// TIA Portal V20 export
FUNCTION_BLOCK "Main_Safety_RTG1"   // FB3, F_LAD
{ S7_Optimized_Access := 'TRUE' }
// stored: AutoNumber false
   VAR
      "ESTOP1_NOT-HALT Taster1" : ESTOP1;
      "stat_Q_NOT-HALT Taster1" : Bool;
      "stat_AckReq_NOT-HALT Taster1" : Bool;
      "ESTOP1_NOT-HALT Extern 1" : ESTOP1;
      "stat_Q_NOT-HALT Extern 1" : Bool;
      "stat_AckReq_NOT-HALT Extern1" : Bool;
      "ESTOP1_NOT-HALT Extern 2" : ESTOP1;
      "stat_Q_NOT-HALT Extern 2" : Bool;
      "stat_AckReq_NOT-HALT Extern 2" : Bool;
      "ESTOP1_Tür 1" : ESTOP1;
      "stat_Q_Tür 1" : Bool;
      "stat_AckReq_Tür 1" : Bool;
      "ESTOP1_Tür 2" : ESTOP1;
      "stat_Q_Tür 2" : Bool;
      "stat_AckReq_Tür 2" : Bool;
      ESTOP1_Systemdruck : ESTOP1;
      stat_AckReq_Systemdruck : Bool;
      "FDBACK_1_NOT-HALT Schütz mit DE_NOT-HALT_Schuetz_Rueckf" : FDBACK;
      "stat_Q_FDBK_1_NOT-HALT Schütz mit DE_NOT-HALT_Schuetz_Rueckf" : Bool;
      "stat_ERROR_FDBK_1_NOT-HALT Schütz mit DE_NOT-HALT_Schuetz_Rueckf" : Bool;
      "FDBACK_2_NOT-HALT Schütz mit IS_Rueck_Entlueftung" : FDBACK;
      "stat_Q_FDBK_2_NOT-HALT Schütz mit IS_Rueck_Entlueftung" : Bool;
      "stat_ERROR_FDBK_2_NOT-HALT Schütz mit IS_Rueck_Entlueftung" : Bool;
      "FDBACK_3_NOT-HALT Schütz mit IS_Druckbereich_entlueftet" : FDBACK;
      "stat_Q_FDBK_3_NOT-HALT Schütz mit IS_Druckbereich_entlueftet" : Bool;
      "stat_ERROR_FDBK_3_NOT-HALT Schütz mit IS_Druckbereich_entlueftet" : Bool;
      "FDBACK_4_NOT-HALT Türe 1 RST mit DE_NOT-HALT_Tuere_1_Rueck_RST" : FDBACK;
      "stat_Q_FDBK_4_NOT-HALT Türe 1 RST mit DE_NOT-HALT_Tuere_1_Rueck_RST" : Bool;
      "stat_ERROR_FDBK_4_NOT-HALT Türe 1 RST mit DE_NOT-HALT_Tuere_1_Rueck_RST" : Bool;
      "FDBACK_5_NOT-HALT Türe 1 mit DE_NOT-HALT_Tuere_1_Rueckf" : FDBACK;
      "stat_Q_FDBK_5_NOT-HALT Türe 1 mit DE_NOT-HALT_Tuere_1_Rueckf" : Bool;
      "stat_ERROR_FDBK_5_NOT-HALT Türe 1 mit DE_NOT-HALT_Tuere_1_Rueckf" : Bool;
      "FDBACK_6_NOT-HALT Türe 1 mit DE_Antriebe_Rueckf" : FDBACK;
      "stat_Q_FDBK_6_NOT-HALT Türe 1 mit DE_Antriebe_Rueckf" : Bool;
      "stat_ERROR_FDBK_6_NOT-HALT Türe 1 mit DE_Antriebe_Rueckf" : Bool;
      "FDBACK_7_NOT-HALT Türe 2 RST mit DE_NOT-HALT_Tuere_2_Rueck_RST" : FDBACK;
      "stat_Q_FDBK_7_NOT-HALT Türe 2 RST mit DE_NOT-HALT_Tuere_2_Rueck_RST" : Bool;
      "stat_ERROR_FDBK_7_NOT-HALT Türe 2 RST mit DE_NOT-HALT_Tuere_2_Rueck_RST" : Bool;
      "FDBACK_8_NOT-HALT Türe 2 mit DE_NOT-HALT_Tuere_2_Rueckf" : FDBACK;
      "stat_Q_FDBK_8_NOT-HALT Türe 2 mit DE_NOT-HALT_Tuere_2_Rueckf" : Bool;
      "stat_ERROR_FDBK_8_NOT-HALT Türe 2 mit DE_NOT-HALT_Tuere_2_Rueckf" : Bool;
      "FDBACK_10_Sicherere Bewegung" : FDBACK;
      "stat_AckReq_10_Sicherere Bewegung" : Bool;
      ACK_GL_Instance : ACK_GL;
      Systemdruck_OK : Bool;
      Antriebe_sicher : Bool;
      "TON_Zuhaltung_Freigben_mit_NOT-HALT" : TON;
      BA_0_groesser_1_5 : Bool;
      TON_BA_0_groesser_1_5 : TON;
      TON_Türen_setzen_zum_öffnen : TON;
      BA_0 : Bool;
      Zuhaltung_freigegeben : Bool;
   END_VAR
BEGIN

REGION Network 1: IS100_0/IS101_0 (2v2) NOT-HALT Taster 1
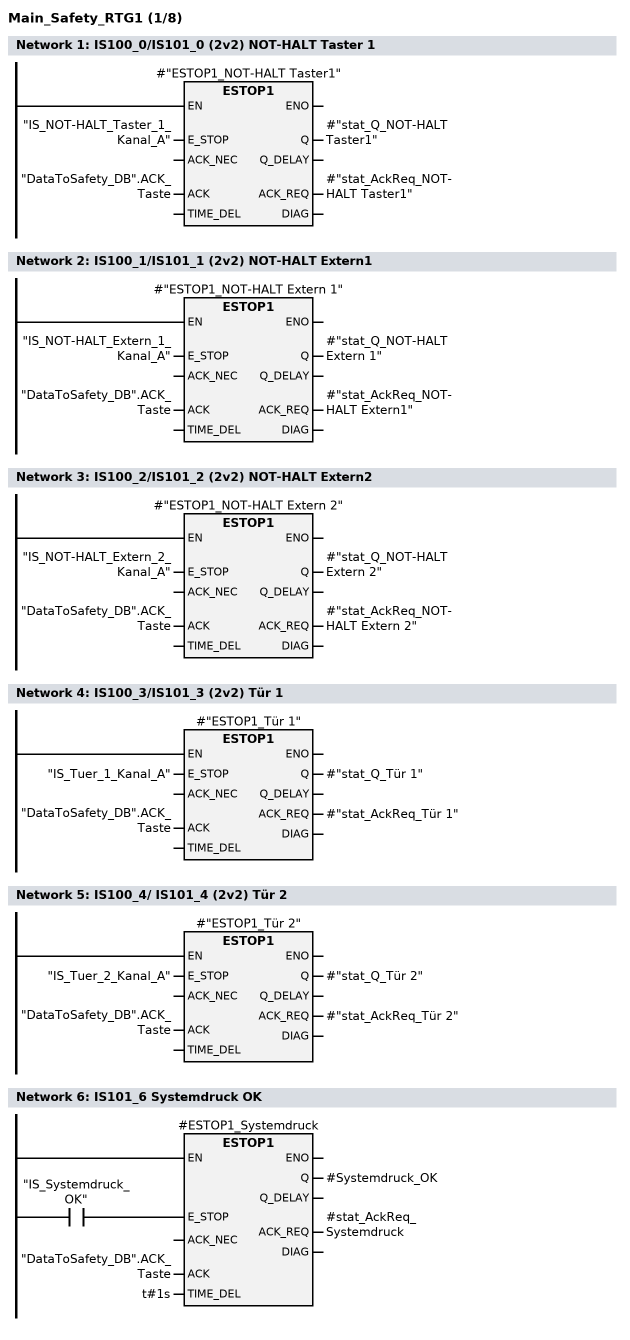
   RUNG wire#powerrail
      #"ESTOP1_NOT-HALT Taster1".ESTOP1(E_STOP := "IS_NOT-HALT_Taster_1_Kanal_A", ACK_NEC :=, ACK := "DataToSafety_DB".ACK_Taste, TIME_DEL :=, Q => #"stat_Q_NOT-HALT Taster1", Q_DELAY =>, ACK_REQ => #"stat_AckReq_NOT-HALT Taster1", DIAG =>)
   END_RUNG
   // the same network as SCL:
   #"ESTOP1_NOT-HALT Taster1"(E_STOP := "IS_NOT-HALT_Taster_1_Kanal_A",   // ESTOP1
                           ACK := "DataToSafety_DB".ACK_Taste,
                           Q => #"stat_Q_NOT-HALT Taster1",
                           ACK_REQ => #"stat_AckReq_NOT-HALT Taster1");
END_REGION

REGION Network 2: IS100_1/IS101_1 (2v2) NOT-HALT Extern1
   RUNG wire#powerrail
      #"ESTOP1_NOT-HALT Extern 1".ESTOP1(E_STOP := "IS_NOT-HALT_Extern_1_Kanal_A", ACK_NEC :=, ACK := "DataToSafety_DB".ACK_Taste, TIME_DEL :=, Q => #"stat_Q_NOT-HALT Extern 1", Q_DELAY =>, ACK_REQ => #"stat_AckReq_NOT-HALT Extern1", DIAG =>)
   END_RUNG
   // the same network as SCL:
   #"ESTOP1_NOT-HALT Extern 1"(E_STOP := "IS_NOT-HALT_Extern_1_Kanal_A",   // ESTOP1
                           ACK := "DataToSafety_DB".ACK_Taste,
                           Q => #"stat_Q_NOT-HALT Extern 1",
                           ACK_REQ => #"stat_AckReq_NOT-HALT Extern1");
END_REGION

REGION Network 3: IS100_2/IS101_2 (2v2) NOT-HALT Extern2
   RUNG wire#powerrail
      #"ESTOP1_NOT-HALT Extern 2".ESTOP1(E_STOP := "IS_NOT-HALT_Extern_2_Kanal_A", ACK_NEC :=, ACK := "DataToSafety_DB".ACK_Taste, TIME_DEL :=, Q => #"stat_Q_NOT-HALT Extern 2", Q_DELAY =>, ACK_REQ => #"stat_AckReq_NOT-HALT Extern 2", DIAG =>)
   END_RUNG
   // the same network as SCL:
   #"ESTOP1_NOT-HALT Extern 2"(E_STOP := "IS_NOT-HALT_Extern_2_Kanal_A",   // ESTOP1
                           ACK := "DataToSafety_DB".ACK_Taste,
                           Q => #"stat_Q_NOT-HALT Extern 2",
                           ACK_REQ => #"stat_AckReq_NOT-HALT Extern 2");
END_REGION

REGION Network 4: IS100_3/IS101_3 (2v2) Tür 1
   RUNG wire#powerrail
      #"ESTOP1_Tür 1".ESTOP1(E_STOP := "IS_Tuer_1_Kanal_A", ACK_NEC :=, ACK := "DataToSafety_DB".ACK_Taste, TIME_DEL :=, Q => #"stat_Q_Tür 1", Q_DELAY =>, ACK_REQ => #"stat_AckReq_Tür 1", DIAG =>)
   END_RUNG
   // the same network as SCL:
   #"ESTOP1_Tür 1"(E_STOP := "IS_Tuer_1_Kanal_A",   // ESTOP1
                   ACK := "DataToSafety_DB".ACK_Taste,
                   Q => #"stat_Q_Tür 1",
                   ACK_REQ => #"stat_AckReq_Tür 1");
END_REGION

REGION Network 5: IS100_4/ IS101_4 (2v2) Tür 2
   RUNG wire#powerrail
      #"ESTOP1_Tür 2".ESTOP1(E_STOP := "IS_Tuer_2_Kanal_A", ACK_NEC :=, ACK := "DataToSafety_DB".ACK_Taste, TIME_DEL :=, Q => #"stat_Q_Tür 2", Q_DELAY =>, ACK_REQ => #"stat_AckReq_Tür 2", DIAG =>)
   END_RUNG
   // the same network as SCL:
   #"ESTOP1_Tür 2"(E_STOP := "IS_Tuer_2_Kanal_A",   // ESTOP1
                   ACK := "DataToSafety_DB".ACK_Taste,
                   Q => #"stat_Q_Tür 2",
                   ACK_REQ => #"stat_AckReq_Tür 2");
END_REGION

REGION Network 6: IS101_6 Systemdruck OK
   RUNG wire#powerrail
      #ESTOP1_Systemdruck.ESTOP1(E_STOP := wire#w1, ACK_NEC :=, ACK := "DataToSafety_DB".ACK_Taste, TIME_DEL := t#1s, Q => #Systemdruck_OK, Q_DELAY =>, ACK_REQ => #stat_AckReq_Systemdruck, DIAG =>)
   END_RUNG
   RUNG wire#powerrail
      Contact( "IS_Systemdruck_OK" )
   END_RUNG wire#w1
   // the same network as SCL:
   #ESTOP1_Systemdruck(E_STOP := "IS_Systemdruck_OK",   // ESTOP1
                       ACK := "DataToSafety_DB".ACK_Taste,
                       TIME_DEL := t#1s,
                       Q => #Systemdruck_OK,
                       ACK_REQ => #stat_AckReq_Systemdruck);
END_REGION

REGION Network 7: Antriebe sicher
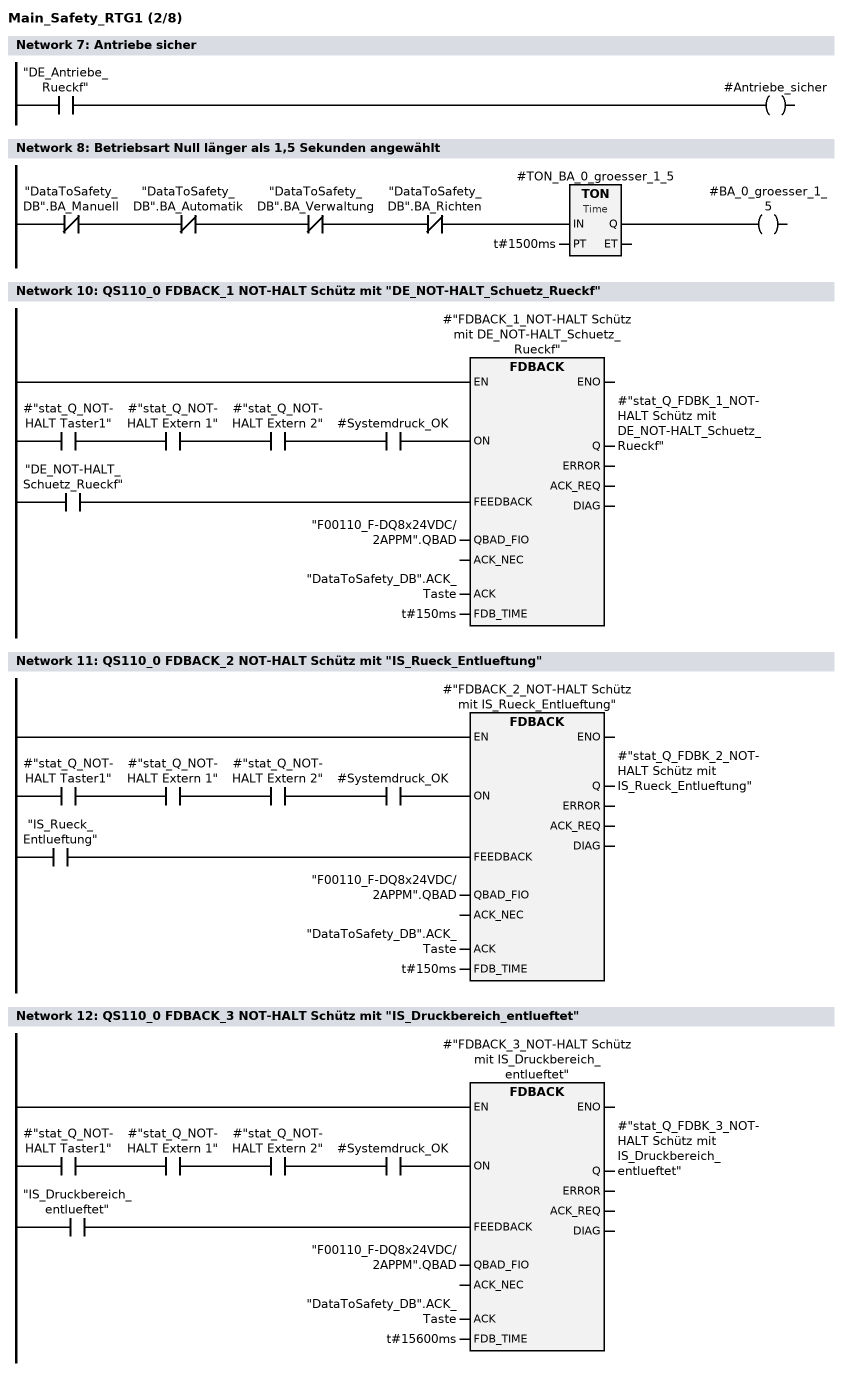
   RUNG wire#powerrail
      Contact( "DE_Antriebe_Rueckf" )
      Coil( #Antriebe_sicher )
   END_RUNG
   // the same network as SCL:
   #Antriebe_sicher := "DE_Antriebe_Rueckf";
END_REGION

REGION Network 8: Betriebsart Null länger als 1,5 Sekunden angewählt
   RUNG wire#powerrail
      I_Contact( "DataToSafety_DB".BA_Manuell )
      I_Contact( "DataToSafety_DB".BA_Automatik )
      I_Contact( "DataToSafety_DB".BA_Verwaltung )
      I_Contact( "DataToSafety_DB".BA_Richten )
      { S7_Templates := "[time_type := Time, codedbool_type := DInt]" } #TON_BA_0_groesser_1_5.TON(pt := t#1500ms, et =>)
      Coil( #BA_0_groesser_1_5 )
   END_RUNG
   // the same network as SCL:
   #TON_BA_0_groesser_1_5.TON(IN := NOT "DataToSafety_DB".BA_Manuell AND NOT "DataToSafety_DB".BA_Automatik AND NOT "DataToSafety_DB".BA_Verwaltung AND NOT "DataToSafety_DB".BA_Richten,
                           PT := t#1500ms);
   #BA_0_groesser_1_5 := #TON_BA_0_groesser_1_5.Q;
END_REGION

REGION Network 9: *********************************************************************************************
END_REGION

REGION Network 10: QS110_0 FDBACK_1 NOT-HALT Schütz mit "DE_NOT-HALT_Schuetz_Rueckf"
   RUNG wire#powerrail
      #"FDBACK_1_NOT-HALT Schütz mit DE_NOT-HALT_Schuetz_Rueckf".FDBACK(ON := wire#w1, FEEDBACK := wire#w2, QBAD_FIO := "F00110_F-DQ8x24VDC/2APPM".QBAD, ACK_NEC :=, ACK := "DataToSafety_DB".ACK_Taste, FDB_TIME := t#150ms, Q => #"stat_Q_FDBK_1_NOT-HALT Schütz mit DE_NOT-HALT_Schuetz_Rueckf", ERROR =>, ACK_REQ =>, DIAG =>)
   END_RUNG
   RUNG wire#powerrail
      Contact( #"stat_Q_NOT-HALT Taster1" )
      Contact( #"stat_Q_NOT-HALT Extern 1" )
      Contact( #"stat_Q_NOT-HALT Extern 2" )
      Contact( #Systemdruck_OK )
   END_RUNG wire#w1
   RUNG wire#powerrail
      Contact( "DE_NOT-HALT_Schuetz_Rueckf" )
   END_RUNG wire#w2
   // the same network as SCL:
   #"FDBACK_1_NOT-HALT Schütz mit DE_NOT-HALT_Schuetz_Rueckf"(ON := #"stat_Q_NOT-HALT Taster1" AND #"stat_Q_NOT-HALT Extern 1" AND #"stat_Q_NOT-HALT Extern 2" AND #Systemdruck_OK,   // FDBACK
                           FEEDBACK := "DE_NOT-HALT_Schuetz_Rueckf",
                           QBAD_FIO := "F00110_F-DQ8x24VDC/2APPM".QBAD,
                           ACK := "DataToSafety_DB".ACK_Taste,
                           FDB_TIME := t#150ms,
                           Q => #"stat_Q_FDBK_1_NOT-HALT Schütz mit DE_NOT-HALT_Schuetz_Rueckf");
END_REGION

REGION Network 11: QS110_0 FDBACK_2 NOT-HALT Schütz mit "IS_Rueck_Entlueftung"
   RUNG wire#powerrail
      #"FDBACK_2_NOT-HALT Schütz mit IS_Rueck_Entlueftung".FDBACK(ON := wire#w1, FEEDBACK := wire#w2, QBAD_FIO := "F00110_F-DQ8x24VDC/2APPM".QBAD, ACK_NEC :=, ACK := "DataToSafety_DB".ACK_Taste, FDB_TIME := t#150ms, Q => #"stat_Q_FDBK_2_NOT-HALT Schütz mit IS_Rueck_Entlueftung", ERROR =>, ACK_REQ =>, DIAG =>)
   END_RUNG
   RUNG wire#powerrail
      Contact( #"stat_Q_NOT-HALT Taster1" )
      Contact( #"stat_Q_NOT-HALT Extern 1" )
      Contact( #"stat_Q_NOT-HALT Extern 2" )
      Contact( #Systemdruck_OK )
   END_RUNG wire#w1
   RUNG wire#powerrail
      Contact( "IS_Rueck_Entlueftung" )
   END_RUNG wire#w2
   // the same network as SCL:
   #"FDBACK_2_NOT-HALT Schütz mit IS_Rueck_Entlueftung"(ON := #"stat_Q_NOT-HALT Taster1" AND #"stat_Q_NOT-HALT Extern 1" AND #"stat_Q_NOT-HALT Extern 2" AND #Systemdruck_OK,   // FDBACK
                           FEEDBACK := "IS_Rueck_Entlueftung",
                           QBAD_FIO := "F00110_F-DQ8x24VDC/2APPM".QBAD,
                           ACK := "DataToSafety_DB".ACK_Taste,
                           FDB_TIME := t#150ms,
                           Q => #"stat_Q_FDBK_2_NOT-HALT Schütz mit IS_Rueck_Entlueftung");
END_REGION

REGION Network 12: QS110_0 FDBACK_3 NOT-HALT Schütz mit "IS_Druckbereich_entlueftet"
   RUNG wire#powerrail
      #"FDBACK_3_NOT-HALT Schütz mit IS_Druckbereich_entlueftet".FDBACK(ON := wire#w1, FEEDBACK := wire#w2, QBAD_FIO := "F00110_F-DQ8x24VDC/2APPM".QBAD, ACK_NEC :=, ACK := "DataToSafety_DB".ACK_Taste, FDB_TIME := t#15600ms, Q => #"stat_Q_FDBK_3_NOT-HALT Schütz mit IS_Druckbereich_entlueftet", ERROR =>, ACK_REQ =>, DIAG =>)
   END_RUNG
   RUNG wire#powerrail
      Contact( #"stat_Q_NOT-HALT Taster1" )
      Contact( #"stat_Q_NOT-HALT Extern 1" )
      Contact( #"stat_Q_NOT-HALT Extern 2" )
      Contact( #Systemdruck_OK )
   END_RUNG wire#w1
   RUNG wire#powerrail
      Contact( "IS_Druckbereich_entlueftet" )
   END_RUNG wire#w2
   // the same network as SCL:
   #"FDBACK_3_NOT-HALT Schütz mit IS_Druckbereich_entlueftet"(ON := #"stat_Q_NOT-HALT Taster1" AND #"stat_Q_NOT-HALT Extern 1" AND #"stat_Q_NOT-HALT Extern 2" AND #Systemdruck_OK,   // FDBACK
                           FEEDBACK := "IS_Druckbereich_entlueftet",
                           QBAD_FIO := "F00110_F-DQ8x24VDC/2APPM".QBAD,
                           ACK := "DataToSafety_DB".ACK_Taste,
                           FDB_TIME := t#15600ms,
                           Q => #"stat_Q_FDBK_3_NOT-HALT Schütz mit IS_Druckbereich_entlueftet");
END_REGION

REGION Network 13: QS110_0 Schütz NOT-HALT Schütz
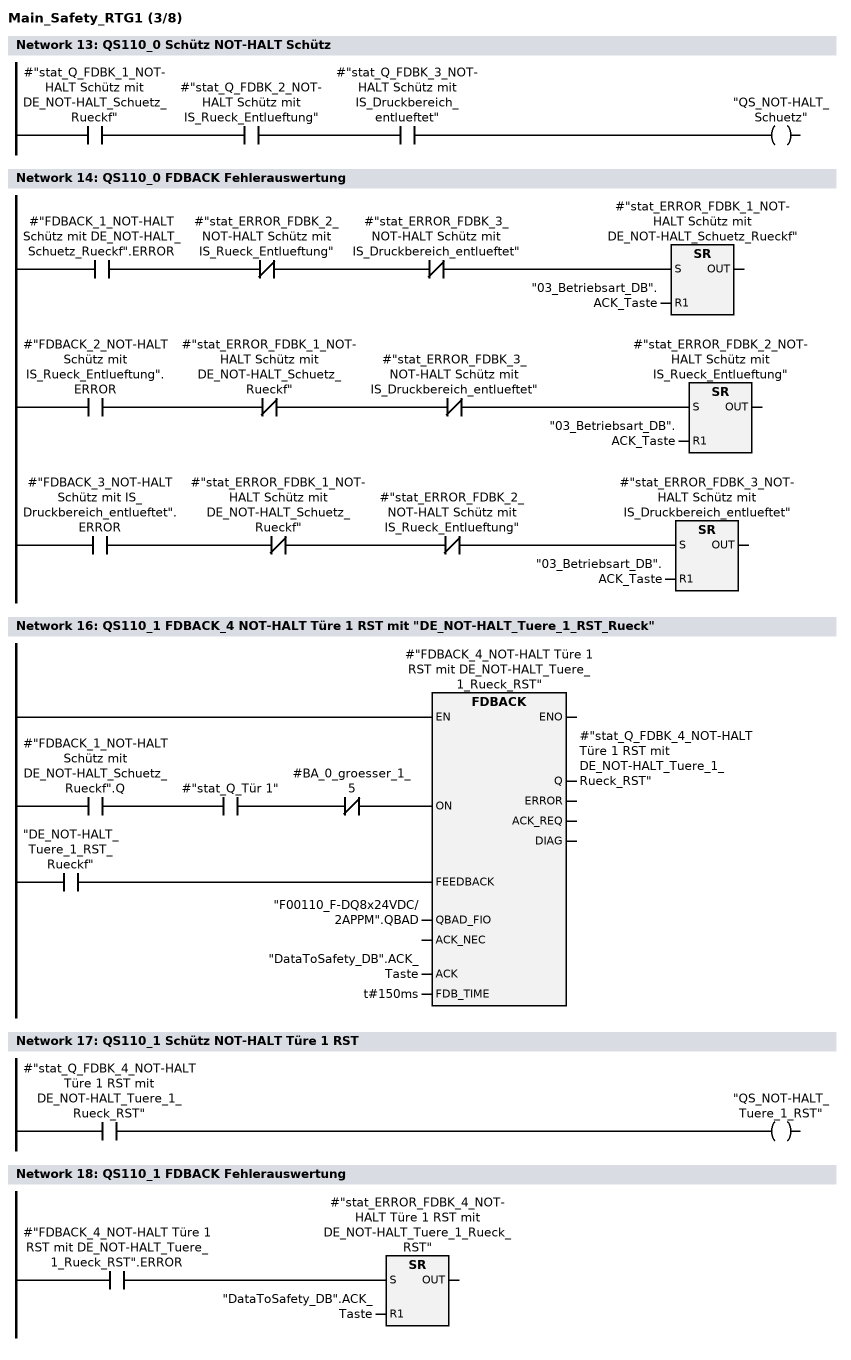
   RUNG wire#powerrail
      Contact( #"stat_Q_FDBK_1_NOT-HALT Schütz mit DE_NOT-HALT_Schuetz_Rueckf" )
      Contact( #"stat_Q_FDBK_2_NOT-HALT Schütz mit IS_Rueck_Entlueftung" )
      Contact( #"stat_Q_FDBK_3_NOT-HALT Schütz mit IS_Druckbereich_entlueftet" )
      Coil( "QS_NOT-HALT_Schuetz" )
   END_RUNG
   // the same network as SCL:
   "QS_NOT-HALT_Schuetz" := #"stat_Q_FDBK_1_NOT-HALT Schütz mit DE_NOT-HALT_Schuetz_Rueckf" AND #"stat_Q_FDBK_2_NOT-HALT Schütz mit IS_Rueck_Entlueftung" AND #"stat_Q_FDBK_3_NOT-HALT Schütz mit IS_Druckbereich_entlueftet";
END_REGION

REGION Network 14: QS110_0 FDBACK Fehlerauswertung
   RUNG wire#powerrail
      Contact( #"FDBACK_1_NOT-HALT Schütz mit DE_NOT-HALT_Schuetz_Rueckf".ERROR )
      I_Contact( #"stat_ERROR_FDBK_2_NOT-HALT Schütz mit IS_Rueck_Entlueftung" )
      I_Contact( #"stat_ERROR_FDBK_3_NOT-HALT Schütz mit IS_Druckbereich_entlueftet" )
      S_SR(operand := #"stat_ERROR_FDBK_1_NOT-HALT Schütz mit DE_NOT-HALT_Schuetz_Rueckf", r1 := "03_Betriebsart_DB".ACK_Taste)
   END_RUNG
   RUNG wire#powerrail
      Contact( #"FDBACK_2_NOT-HALT Schütz mit IS_Rueck_Entlueftung".ERROR )
      I_Contact( #"stat_ERROR_FDBK_1_NOT-HALT Schütz mit DE_NOT-HALT_Schuetz_Rueckf" )
      I_Contact( #"stat_ERROR_FDBK_3_NOT-HALT Schütz mit IS_Druckbereich_entlueftet" )
      S_SR(operand := #"stat_ERROR_FDBK_2_NOT-HALT Schütz mit IS_Rueck_Entlueftung", r1 := "03_Betriebsart_DB".ACK_Taste)
   END_RUNG
   RUNG wire#powerrail
      Contact( #"FDBACK_3_NOT-HALT Schütz mit IS_Druckbereich_entlueftet".ERROR )
      I_Contact( #"stat_ERROR_FDBK_1_NOT-HALT Schütz mit DE_NOT-HALT_Schuetz_Rueckf" )
      I_Contact( #"stat_ERROR_FDBK_2_NOT-HALT Schütz mit IS_Rueck_Entlueftung" )
      S_SR(operand := #"stat_ERROR_FDBK_3_NOT-HALT Schütz mit IS_Druckbereich_entlueftet", r1 := "03_Betriebsart_DB".ACK_Taste)
   END_RUNG
   // the same network as SCL:
   IF #"FDBACK_1_NOT-HALT Schütz mit DE_NOT-HALT_Schuetz_Rueckf".ERROR AND NOT #"stat_ERROR_FDBK_2_NOT-HALT Schütz mit IS_Rueck_Entlueftung" AND NOT #"stat_ERROR_FDBK_3_NOT-HALT Schütz mit IS_Druckbereich_entlueftet" THEN
       #"stat_ERROR_FDBK_1_NOT-HALT Schütz mit DE_NOT-HALT_Schuetz_Rueckf" := TRUE;   // SR flip-flop
   END_IF;
   IF "03_Betriebsart_DB".ACK_Taste THEN
       #"stat_ERROR_FDBK_1_NOT-HALT Schütz mit DE_NOT-HALT_Schuetz_Rueckf" := FALSE;
   END_IF;
   IF #"FDBACK_2_NOT-HALT Schütz mit IS_Rueck_Entlueftung".ERROR AND NOT #"stat_ERROR_FDBK_1_NOT-HALT Schütz mit DE_NOT-HALT_Schuetz_Rueckf" AND NOT #"stat_ERROR_FDBK_3_NOT-HALT Schütz mit IS_Druckbereich_entlueftet" THEN
       #"stat_ERROR_FDBK_2_NOT-HALT Schütz mit IS_Rueck_Entlueftung" := TRUE;   // SR flip-flop
   END_IF;
   IF "03_Betriebsart_DB".ACK_Taste THEN
       #"stat_ERROR_FDBK_2_NOT-HALT Schütz mit IS_Rueck_Entlueftung" := FALSE;
   END_IF;
   IF #"FDBACK_3_NOT-HALT Schütz mit IS_Druckbereich_entlueftet".ERROR AND NOT #"stat_ERROR_FDBK_1_NOT-HALT Schütz mit DE_NOT-HALT_Schuetz_Rueckf" AND NOT #"stat_ERROR_FDBK_2_NOT-HALT Schütz mit IS_Rueck_Entlueftung" THEN
       #"stat_ERROR_FDBK_3_NOT-HALT Schütz mit IS_Druckbereich_entlueftet" := TRUE;   // SR flip-flop
   END_IF;
   IF "03_Betriebsart_DB".ACK_Taste THEN
       #"stat_ERROR_FDBK_3_NOT-HALT Schütz mit IS_Druckbereich_entlueftet" := FALSE;
   END_IF;
END_REGION

REGION Network 15: *********************************************************************************************
END_REGION

REGION Network 16: QS110_1 FDBACK_4 NOT-HALT Türe 1 RST mit "DE_NOT-HALT_Tuere_1_RST_Rueck"
   RUNG wire#powerrail
      #"FDBACK_4_NOT-HALT Türe 1 RST mit DE_NOT-HALT_Tuere_1_Rueck_RST".FDBACK(ON := wire#w1, FEEDBACK := wire#w2, QBAD_FIO := "F00110_F-DQ8x24VDC/2APPM".QBAD, ACK_NEC :=, ACK := "DataToSafety_DB".ACK_Taste, FDB_TIME := t#150ms, Q => #"stat_Q_FDBK_4_NOT-HALT Türe 1 RST mit DE_NOT-HALT_Tuere_1_Rueck_RST", ERROR =>, ACK_REQ =>, DIAG =>)
   END_RUNG
   RUNG wire#powerrail
      Contact( #"FDBACK_1_NOT-HALT Schütz mit DE_NOT-HALT_Schuetz_Rueckf".Q )
      Contact( #"stat_Q_Tür 1" )
      I_Contact( #BA_0_groesser_1_5 )
   END_RUNG wire#w1
   RUNG wire#powerrail
      Contact( "DE_NOT-HALT_Tuere_1_RST_Rueckf" )
   END_RUNG wire#w2
   // the same network as SCL:
   #"FDBACK_4_NOT-HALT Türe 1 RST mit DE_NOT-HALT_Tuere_1_Rueck_RST"(ON := #"FDBACK_1_NOT-HALT Schütz mit DE_NOT-HALT_Schuetz_Rueckf".Q AND #"stat_Q_Tür 1" AND NOT #BA_0_groesser_1_5,   // FDBACK
                           FEEDBACK := "DE_NOT-HALT_Tuere_1_RST_Rueckf",
                           QBAD_FIO := "F00110_F-DQ8x24VDC/2APPM".QBAD,
                           ACK := "DataToSafety_DB".ACK_Taste,
                           FDB_TIME := t#150ms,
                           Q => #"stat_Q_FDBK_4_NOT-HALT Türe 1 RST mit DE_NOT-HALT_Tuere_1_Rueck_RST");
END_REGION

REGION Network 17: QS110_1 Schütz NOT-HALT Türe 1 RST
   RUNG wire#powerrail
      Contact( #"stat_Q_FDBK_4_NOT-HALT Türe 1 RST mit DE_NOT-HALT_Tuere_1_Rueck_RST" )
      Coil( "QS_NOT-HALT_Tuere_1_RST" )
   END_RUNG
   // the same network as SCL:
   "QS_NOT-HALT_Tuere_1_RST" := #"stat_Q_FDBK_4_NOT-HALT Türe 1 RST mit DE_NOT-HALT_Tuere_1_Rueck_RST";
END_REGION

REGION Network 18: QS110_1 FDBACK Fehlerauswertung
   RUNG wire#powerrail
      Contact( #"FDBACK_4_NOT-HALT Türe 1 RST mit DE_NOT-HALT_Tuere_1_Rueck_RST".ERROR )
      S_SR(operand := #"stat_ERROR_FDBK_4_NOT-HALT Türe 1 RST mit DE_NOT-HALT_Tuere_1_Rueck_RST", r1 := "DataToSafety_DB".ACK_Taste)
   END_RUNG
   // the same network as SCL:
   IF #"FDBACK_4_NOT-HALT Türe 1 RST mit DE_NOT-HALT_Tuere_1_Rueck_RST".ERROR THEN
       #"stat_ERROR_FDBK_4_NOT-HALT Türe 1 RST mit DE_NOT-HALT_Tuere_1_Rueck_RST" := TRUE;   // SR flip-flop
   END_IF;
   IF "DataToSafety_DB".ACK_Taste THEN
       #"stat_ERROR_FDBK_4_NOT-HALT Türe 1 RST mit DE_NOT-HALT_Tuere_1_Rueck_RST" := FALSE;
   END_IF;
END_REGION

REGION Network 19: *********************************************************************************************
END_REGION

REGION Network 20: QS110_2 FDBACK_5 NOT-HALT Türe 1 mit "DE_NOT-HALT_Tuere_1_Rueckf"
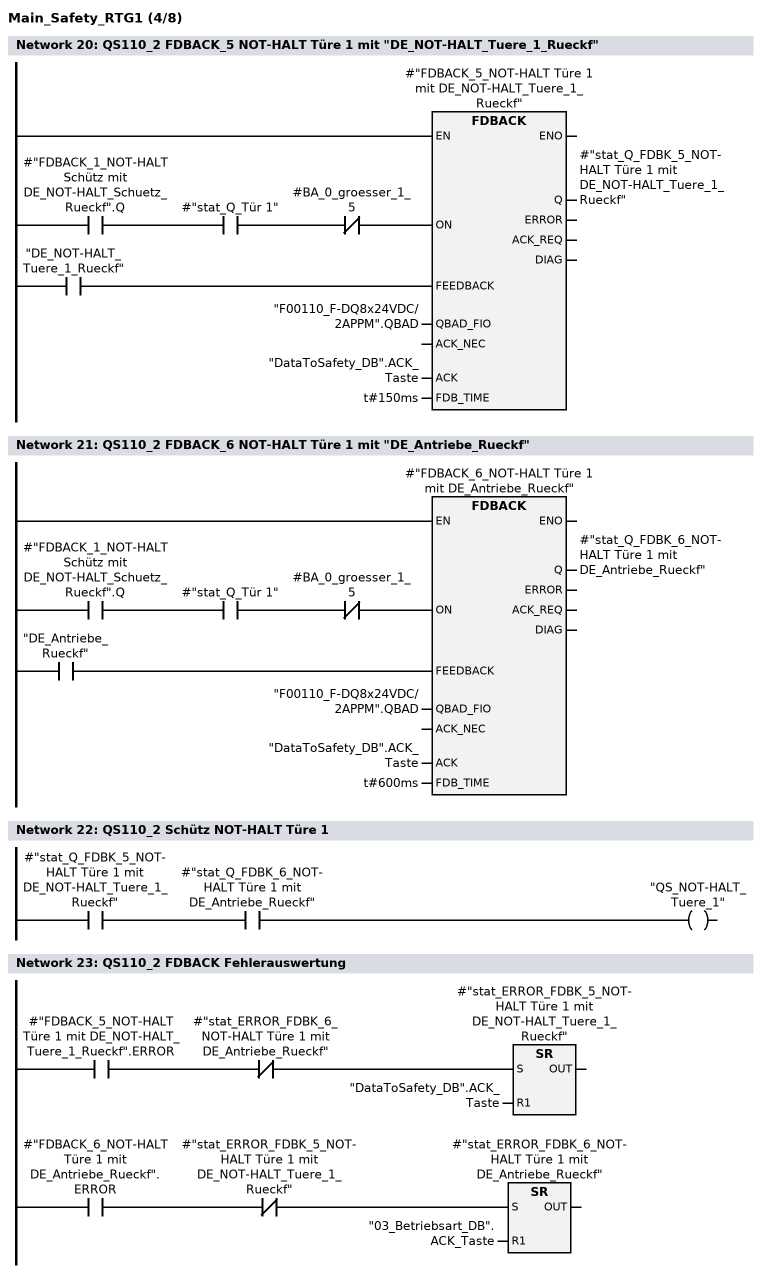
   RUNG wire#powerrail
      #"FDBACK_5_NOT-HALT Türe 1 mit DE_NOT-HALT_Tuere_1_Rueckf".FDBACK(ON := wire#w1, FEEDBACK := wire#w2, QBAD_FIO := "F00110_F-DQ8x24VDC/2APPM".QBAD, ACK_NEC :=, ACK := "DataToSafety_DB".ACK_Taste, FDB_TIME := t#150ms, Q => #"stat_Q_FDBK_5_NOT-HALT Türe 1 mit DE_NOT-HALT_Tuere_1_Rueckf", ERROR =>, ACK_REQ =>, DIAG =>)
   END_RUNG
   RUNG wire#powerrail
      Contact( #"FDBACK_1_NOT-HALT Schütz mit DE_NOT-HALT_Schuetz_Rueckf".Q )
      Contact( #"stat_Q_Tür 1" )
      I_Contact( #BA_0_groesser_1_5 )
   END_RUNG wire#w1
   RUNG wire#powerrail
      Contact( "DE_NOT-HALT_Tuere_1_Rueckf" )
   END_RUNG wire#w2
   // the same network as SCL:
   #"FDBACK_5_NOT-HALT Türe 1 mit DE_NOT-HALT_Tuere_1_Rueckf"(ON := #"FDBACK_1_NOT-HALT Schütz mit DE_NOT-HALT_Schuetz_Rueckf".Q AND #"stat_Q_Tür 1" AND NOT #BA_0_groesser_1_5,   // FDBACK
                           FEEDBACK := "DE_NOT-HALT_Tuere_1_Rueckf",
                           QBAD_FIO := "F00110_F-DQ8x24VDC/2APPM".QBAD,
                           ACK := "DataToSafety_DB".ACK_Taste,
                           FDB_TIME := t#150ms,
                           Q => #"stat_Q_FDBK_5_NOT-HALT Türe 1 mit DE_NOT-HALT_Tuere_1_Rueckf");
END_REGION

REGION Network 21: QS110_2 FDBACK_6 NOT-HALT Türe 1 mit "DE_Antriebe_Rueckf"
   RUNG wire#powerrail
      #"FDBACK_6_NOT-HALT Türe 1 mit DE_Antriebe_Rueckf".FDBACK(ON := wire#w1, FEEDBACK := wire#w2, QBAD_FIO := "F00110_F-DQ8x24VDC/2APPM".QBAD, ACK_NEC :=, ACK := "DataToSafety_DB".ACK_Taste, FDB_TIME := t#600ms, Q => #"stat_Q_FDBK_6_NOT-HALT Türe 1 mit DE_Antriebe_Rueckf", ERROR =>, ACK_REQ =>, DIAG =>)
   END_RUNG
   RUNG wire#powerrail
      Contact( #"FDBACK_1_NOT-HALT Schütz mit DE_NOT-HALT_Schuetz_Rueckf".Q )
      Contact( #"stat_Q_Tür 1" )
      I_Contact( #BA_0_groesser_1_5 )
   END_RUNG wire#w1
   RUNG wire#powerrail
      Contact( "DE_Antriebe_Rueckf" )
   END_RUNG wire#w2
   // the same network as SCL:
   #"FDBACK_6_NOT-HALT Türe 1 mit DE_Antriebe_Rueckf"(ON := #"FDBACK_1_NOT-HALT Schütz mit DE_NOT-HALT_Schuetz_Rueckf".Q AND #"stat_Q_Tür 1" AND NOT #BA_0_groesser_1_5,   // FDBACK
                           FEEDBACK := "DE_Antriebe_Rueckf",
                           QBAD_FIO := "F00110_F-DQ8x24VDC/2APPM".QBAD,
                           ACK := "DataToSafety_DB".ACK_Taste,
                           FDB_TIME := t#600ms,
                           Q => #"stat_Q_FDBK_6_NOT-HALT Türe 1 mit DE_Antriebe_Rueckf");
END_REGION

REGION Network 22: QS110_2 Schütz NOT-HALT Türe 1
   RUNG wire#powerrail
      Contact( #"stat_Q_FDBK_5_NOT-HALT Türe 1 mit DE_NOT-HALT_Tuere_1_Rueckf" )
      Contact( #"stat_Q_FDBK_6_NOT-HALT Türe 1 mit DE_Antriebe_Rueckf" )
      Coil( "QS_NOT-HALT_Tuere_1" )
   END_RUNG
   // the same network as SCL:
   "QS_NOT-HALT_Tuere_1" := #"stat_Q_FDBK_5_NOT-HALT Türe 1 mit DE_NOT-HALT_Tuere_1_Rueckf" AND #"stat_Q_FDBK_6_NOT-HALT Türe 1 mit DE_Antriebe_Rueckf";
END_REGION

REGION Network 23: QS110_2 FDBACK Fehlerauswertung
   RUNG wire#powerrail
      Contact( #"FDBACK_5_NOT-HALT Türe 1 mit DE_NOT-HALT_Tuere_1_Rueckf".ERROR )
      I_Contact( #"stat_ERROR_FDBK_6_NOT-HALT Türe 1 mit DE_Antriebe_Rueckf" )
      S_SR(operand := #"stat_ERROR_FDBK_5_NOT-HALT Türe 1 mit DE_NOT-HALT_Tuere_1_Rueckf", r1 := "DataToSafety_DB".ACK_Taste)
   END_RUNG
   RUNG wire#powerrail
      Contact( #"FDBACK_6_NOT-HALT Türe 1 mit DE_Antriebe_Rueckf".ERROR )
      I_Contact( #"stat_ERROR_FDBK_5_NOT-HALT Türe 1 mit DE_NOT-HALT_Tuere_1_Rueckf" )
      S_SR(operand := #"stat_ERROR_FDBK_6_NOT-HALT Türe 1 mit DE_Antriebe_Rueckf", r1 := "03_Betriebsart_DB".ACK_Taste)
   END_RUNG
   // the same network as SCL:
   IF #"FDBACK_5_NOT-HALT Türe 1 mit DE_NOT-HALT_Tuere_1_Rueckf".ERROR AND NOT #"stat_ERROR_FDBK_6_NOT-HALT Türe 1 mit DE_Antriebe_Rueckf" THEN
       #"stat_ERROR_FDBK_5_NOT-HALT Türe 1 mit DE_NOT-HALT_Tuere_1_Rueckf" := TRUE;   // SR flip-flop
   END_IF;
   IF "DataToSafety_DB".ACK_Taste THEN
       #"stat_ERROR_FDBK_5_NOT-HALT Türe 1 mit DE_NOT-HALT_Tuere_1_Rueckf" := FALSE;
   END_IF;
   IF #"FDBACK_6_NOT-HALT Türe 1 mit DE_Antriebe_Rueckf".ERROR AND NOT #"stat_ERROR_FDBK_5_NOT-HALT Türe 1 mit DE_NOT-HALT_Tuere_1_Rueckf" THEN
       #"stat_ERROR_FDBK_6_NOT-HALT Türe 1 mit DE_Antriebe_Rueckf" := TRUE;   // SR flip-flop
   END_IF;
   IF "03_Betriebsart_DB".ACK_Taste THEN
       #"stat_ERROR_FDBK_6_NOT-HALT Türe 1 mit DE_Antriebe_Rueckf" := FALSE;
   END_IF;
END_REGION

REGION Network 24: *********************************************************************************************
END_REGION

REGION Network 25: QS110_3 FDBACK_7 NOT-HALT Türe 2 RST mit "DE_NOT-HALT_Tuere_2_RST_Rueck"
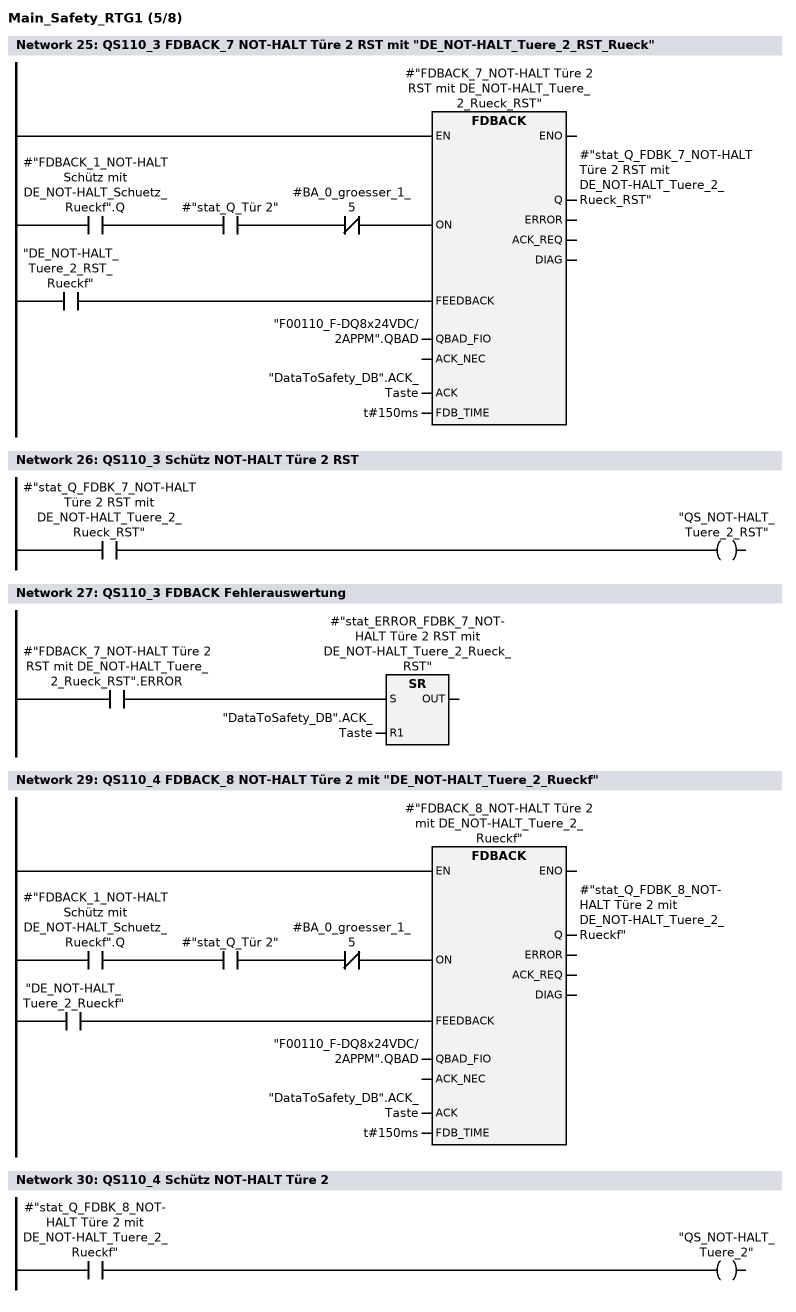
   RUNG wire#powerrail
      #"FDBACK_7_NOT-HALT Türe 2 RST mit DE_NOT-HALT_Tuere_2_Rueck_RST".FDBACK(ON := wire#w1, FEEDBACK := wire#w2, QBAD_FIO := "F00110_F-DQ8x24VDC/2APPM".QBAD, ACK_NEC :=, ACK := "DataToSafety_DB".ACK_Taste, FDB_TIME := t#150ms, Q => #"stat_Q_FDBK_7_NOT-HALT Türe 2 RST mit DE_NOT-HALT_Tuere_2_Rueck_RST", ERROR =>, ACK_REQ =>, DIAG =>)
   END_RUNG
   RUNG wire#powerrail
      Contact( #"FDBACK_1_NOT-HALT Schütz mit DE_NOT-HALT_Schuetz_Rueckf".Q )
      Contact( #"stat_Q_Tür 2" )
      I_Contact( #BA_0_groesser_1_5 )
   END_RUNG wire#w1
   RUNG wire#powerrail
      Contact( "DE_NOT-HALT_Tuere_2_RST_Rueckf" )
   END_RUNG wire#w2
   // the same network as SCL:
   #"FDBACK_7_NOT-HALT Türe 2 RST mit DE_NOT-HALT_Tuere_2_Rueck_RST"(ON := #"FDBACK_1_NOT-HALT Schütz mit DE_NOT-HALT_Schuetz_Rueckf".Q AND #"stat_Q_Tür 2" AND NOT #BA_0_groesser_1_5,   // FDBACK
                           FEEDBACK := "DE_NOT-HALT_Tuere_2_RST_Rueckf",
                           QBAD_FIO := "F00110_F-DQ8x24VDC/2APPM".QBAD,
                           ACK := "DataToSafety_DB".ACK_Taste,
                           FDB_TIME := t#150ms,
                           Q => #"stat_Q_FDBK_7_NOT-HALT Türe 2 RST mit DE_NOT-HALT_Tuere_2_Rueck_RST");
END_REGION

REGION Network 26: QS110_3 Schütz NOT-HALT Türe 2 RST
   RUNG wire#powerrail
      Contact( #"stat_Q_FDBK_7_NOT-HALT Türe 2 RST mit DE_NOT-HALT_Tuere_2_Rueck_RST" )
      Coil( "QS_NOT-HALT_Tuere_2_RST" )
   END_RUNG
   // the same network as SCL:
   "QS_NOT-HALT_Tuere_2_RST" := #"stat_Q_FDBK_7_NOT-HALT Türe 2 RST mit DE_NOT-HALT_Tuere_2_Rueck_RST";
END_REGION

REGION Network 27: QS110_3 FDBACK Fehlerauswertung
   RUNG wire#powerrail
      Contact( #"FDBACK_7_NOT-HALT Türe 2 RST mit DE_NOT-HALT_Tuere_2_Rueck_RST".ERROR )
      S_SR(operand := #"stat_ERROR_FDBK_7_NOT-HALT Türe 2 RST mit DE_NOT-HALT_Tuere_2_Rueck_RST", r1 := "DataToSafety_DB".ACK_Taste)
   END_RUNG
   // the same network as SCL:
   IF #"FDBACK_7_NOT-HALT Türe 2 RST mit DE_NOT-HALT_Tuere_2_Rueck_RST".ERROR THEN
       #"stat_ERROR_FDBK_7_NOT-HALT Türe 2 RST mit DE_NOT-HALT_Tuere_2_Rueck_RST" := TRUE;   // SR flip-flop
   END_IF;
   IF "DataToSafety_DB".ACK_Taste THEN
       #"stat_ERROR_FDBK_7_NOT-HALT Türe 2 RST mit DE_NOT-HALT_Tuere_2_Rueck_RST" := FALSE;
   END_IF;
END_REGION

REGION Network 28: *********************************************************************************************
END_REGION

REGION Network 29: QS110_4 FDBACK_8 NOT-HALT Türe 2 mit "DE_NOT-HALT_Tuere_2_Rueckf"
   RUNG wire#powerrail
      #"FDBACK_8_NOT-HALT Türe 2 mit DE_NOT-HALT_Tuere_2_Rueckf".FDBACK(ON := wire#w1, FEEDBACK := wire#w2, QBAD_FIO := "F00110_F-DQ8x24VDC/2APPM".QBAD, ACK_NEC :=, ACK := "DataToSafety_DB".ACK_Taste, FDB_TIME := t#150ms, Q => #"stat_Q_FDBK_8_NOT-HALT Türe 2 mit DE_NOT-HALT_Tuere_2_Rueckf", ERROR =>, ACK_REQ =>, DIAG =>)
   END_RUNG
   RUNG wire#powerrail
      Contact( #"FDBACK_1_NOT-HALT Schütz mit DE_NOT-HALT_Schuetz_Rueckf".Q )
      Contact( #"stat_Q_Tür 2" )
      I_Contact( #BA_0_groesser_1_5 )
   END_RUNG wire#w1
   RUNG wire#powerrail
      Contact( "DE_NOT-HALT_Tuere_2_Rueckf" )
   END_RUNG wire#w2
   // the same network as SCL:
   #"FDBACK_8_NOT-HALT Türe 2 mit DE_NOT-HALT_Tuere_2_Rueckf"(ON := #"FDBACK_1_NOT-HALT Schütz mit DE_NOT-HALT_Schuetz_Rueckf".Q AND #"stat_Q_Tür 2" AND NOT #BA_0_groesser_1_5,   // FDBACK
                           FEEDBACK := "DE_NOT-HALT_Tuere_2_Rueckf",
                           QBAD_FIO := "F00110_F-DQ8x24VDC/2APPM".QBAD,
                           ACK := "DataToSafety_DB".ACK_Taste,
                           FDB_TIME := t#150ms,
                           Q => #"stat_Q_FDBK_8_NOT-HALT Türe 2 mit DE_NOT-HALT_Tuere_2_Rueckf");
END_REGION

REGION Network 30: QS110_4 Schütz NOT-HALT Türe 2
   RUNG wire#powerrail
      Contact( #"stat_Q_FDBK_8_NOT-HALT Türe 2 mit DE_NOT-HALT_Tuere_2_Rueckf" )
      Coil( "QS_NOT-HALT_Tuere_2" )
   END_RUNG
   // the same network as SCL:
   "QS_NOT-HALT_Tuere_2" := #"stat_Q_FDBK_8_NOT-HALT Türe 2 mit DE_NOT-HALT_Tuere_2_Rueckf";
END_REGION

REGION Network 31: QS110_4 FDBACK Fehlerauswertung
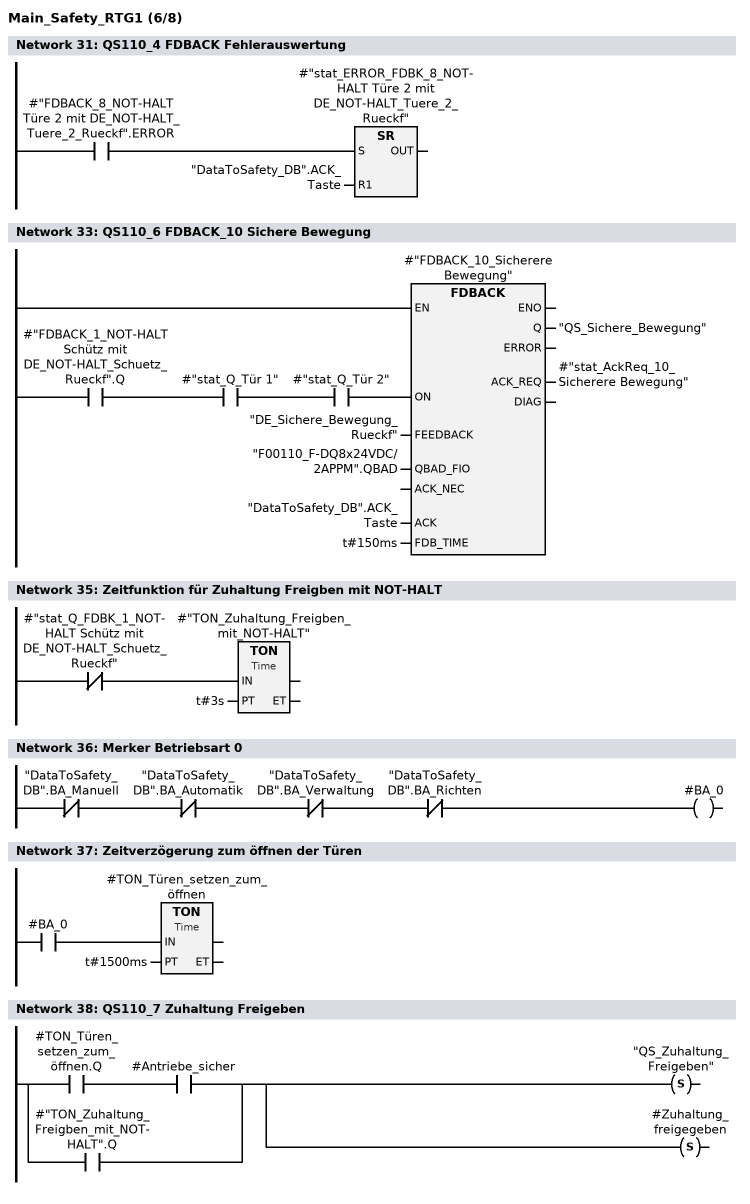
   RUNG wire#powerrail
      Contact( #"FDBACK_8_NOT-HALT Türe 2 mit DE_NOT-HALT_Tuere_2_Rueckf".ERROR )
      S_SR(operand := #"stat_ERROR_FDBK_8_NOT-HALT Türe 2 mit DE_NOT-HALT_Tuere_2_Rueckf", r1 := "DataToSafety_DB".ACK_Taste)
   END_RUNG
   // the same network as SCL:
   IF #"FDBACK_8_NOT-HALT Türe 2 mit DE_NOT-HALT_Tuere_2_Rueckf".ERROR THEN
       #"stat_ERROR_FDBK_8_NOT-HALT Türe 2 mit DE_NOT-HALT_Tuere_2_Rueckf" := TRUE;   // SR flip-flop
   END_IF;
   IF "DataToSafety_DB".ACK_Taste THEN
       #"stat_ERROR_FDBK_8_NOT-HALT Türe 2 mit DE_NOT-HALT_Tuere_2_Rueckf" := FALSE;
   END_IF;
END_REGION

REGION Network 32: *********************************************************************************************
END_REGION

REGION Network 33: QS110_6 FDBACK_10 Sichere Bewegung
   RUNG wire#powerrail
      #"FDBACK_10_Sicherere Bewegung".FDBACK(ON := wire#w1, FEEDBACK := "DE_Sichere_Bewegung_Rueckf", QBAD_FIO := "F00110_F-DQ8x24VDC/2APPM".QBAD, ACK_NEC :=, ACK := "DataToSafety_DB".ACK_Taste, FDB_TIME := t#150ms, Q => "QS_Sichere_Bewegung", ERROR =>, ACK_REQ => #"stat_AckReq_10_Sicherere Bewegung", DIAG =>)
   END_RUNG
   RUNG wire#powerrail
      Contact( #"FDBACK_1_NOT-HALT Schütz mit DE_NOT-HALT_Schuetz_Rueckf".Q )
      Contact( #"stat_Q_Tür 1" )
      Contact( #"stat_Q_Tür 2" )
   END_RUNG wire#w1
   // the same network as SCL:
   #"FDBACK_10_Sicherere Bewegung"(ON := #"FDBACK_1_NOT-HALT Schütz mit DE_NOT-HALT_Schuetz_Rueckf".Q AND #"stat_Q_Tür 1" AND #"stat_Q_Tür 2",   // FDBACK
                           FEEDBACK := "DE_Sichere_Bewegung_Rueckf",
                           QBAD_FIO := "F00110_F-DQ8x24VDC/2APPM".QBAD,
                           ACK := "DataToSafety_DB".ACK_Taste,
                           FDB_TIME := t#150ms,
                           Q => "QS_Sichere_Bewegung",
                           ACK_REQ => #"stat_AckReq_10_Sicherere Bewegung");
END_REGION

REGION Network 34: *********************************************************************************************
END_REGION

REGION Network 35: Zeitfunktion für Zuhaltung Freigben mit NOT-HALT
   RUNG wire#powerrail
      I_Contact( #"stat_Q_FDBK_1_NOT-HALT Schütz mit DE_NOT-HALT_Schuetz_Rueckf" )
      { S7_Templates := "[time_type := Time, codedbool_type := DInt]" } #"TON_Zuhaltung_Freigben_mit_NOT-HALT".TON(pt := t#3s, et =>)
   END_RUNG
   // the same network as SCL:
   #"TON_Zuhaltung_Freigben_mit_NOT-HALT".TON(IN := NOT #"stat_Q_FDBK_1_NOT-HALT Schütz mit DE_NOT-HALT_Schuetz_Rueckf",
                           PT := t#3s);
END_REGION

REGION Network 36: Merker Betriebsart 0
   RUNG wire#powerrail
      I_Contact( "DataToSafety_DB".BA_Manuell )
      I_Contact( "DataToSafety_DB".BA_Automatik )
      I_Contact( "DataToSafety_DB".BA_Verwaltung )
      I_Contact( "DataToSafety_DB".BA_Richten )
      Coil( #BA_0 )
   END_RUNG
   // the same network as SCL:
   #BA_0 := NOT "DataToSafety_DB".BA_Manuell AND NOT "DataToSafety_DB".BA_Automatik AND NOT "DataToSafety_DB".BA_Verwaltung AND NOT "DataToSafety_DB".BA_Richten;
END_REGION

REGION Network 37: Zeitverzögerung zum öffnen der Türen
   RUNG wire#powerrail
      Contact( #BA_0 )
      { S7_Templates := "[time_type := Time, codedbool_type := DInt]" } #TON_Türen_setzen_zum_öffnen.TON(pt := t#1500ms, et =>)
   END_RUNG
   // the same network as SCL:
   #TON_Türen_setzen_zum_öffnen.TON(IN := #BA_0, PT := t#1500ms);
END_REGION

REGION Network 38: QS110_7 Zuhaltung Freigeben
   RUNG wire#powerrail
      Contact( #TON_Türen_setzen_zum_öffnen.Q )
      Contact( #Antriebe_sicher )
      wire#w1
      S_Coil( "QS_Zuhaltung_Freigeben" )
   END_RUNG
   RUNG wire#powerrail
      Contact( #"TON_Zuhaltung_Freigben_mit_NOT-HALT".Q )
   END_RUNG wire#w1
   RUNG wire#w1
      S_Coil( #Zuhaltung_freigegeben )
   END_RUNG
   // the same network as SCL:
   IF (#TON_Türen_setzen_zum_öffnen.Q AND #Antriebe_sicher) OR #"TON_Zuhaltung_Freigben_mit_NOT-HALT".Q THEN
       "QS_Zuhaltung_Freigeben" := TRUE;
       #Zuhaltung_freigegeben := TRUE;
   END_IF;
END_REGION

REGION Network 39: QS110_7 Zuhaltung verriegeln zum schliessen
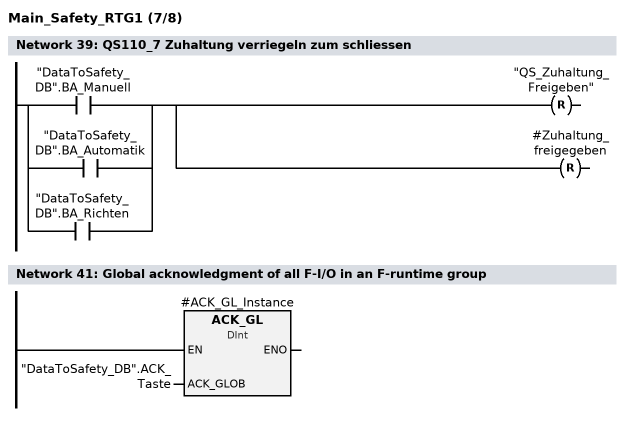
   RUNG wire#powerrail
      Contact( "DataToSafety_DB".BA_Manuell )
      wire#w1
      R_Coil( "QS_Zuhaltung_Freigeben" )
   END_RUNG
   RUNG wire#powerrail
      Contact( "DataToSafety_DB".BA_Automatik )
   END_RUNG wire#w1
   RUNG wire#powerrail
      Contact( "DataToSafety_DB".BA_Richten )
   END_RUNG wire#w1
   RUNG wire#w1
      R_Coil( #Zuhaltung_freigegeben )
   END_RUNG
   // the same network as SCL:
   IF "DataToSafety_DB".BA_Manuell OR "DataToSafety_DB".BA_Automatik OR "DataToSafety_DB".BA_Richten THEN
       "QS_Zuhaltung_Freigeben" := FALSE;
       #Zuhaltung_freigegeben := FALSE;
   END_IF;
END_REGION

REGION Network 40: *********************************************************************************************
END_REGION

REGION Network 41: Global acknowledgment of all F-I/O in an F-runtime group
   RUNG wire#powerrail
      { S7_Templates := "codedbool_type := DInt" } #ACK_GL_Instance.ACK_GL(ACK_GLOB := "DataToSafety_DB".ACK_Taste)
   END_RUNG
   // the same network as SCL:
   #ACK_GL_Instance(ACK_GLOB := "DataToSafety_DB".ACK_Taste);   // ACK_GL
END_REGION

REGION Network 42: Daten von Safety-SPS zur Standard SPS
   // Dieses Netzwerk sammelt mögliche Fehler im Sicherheitsprogramm und schreibt sie in den Datenbaustein um Daten an das Standardprogramm zu übergeben.
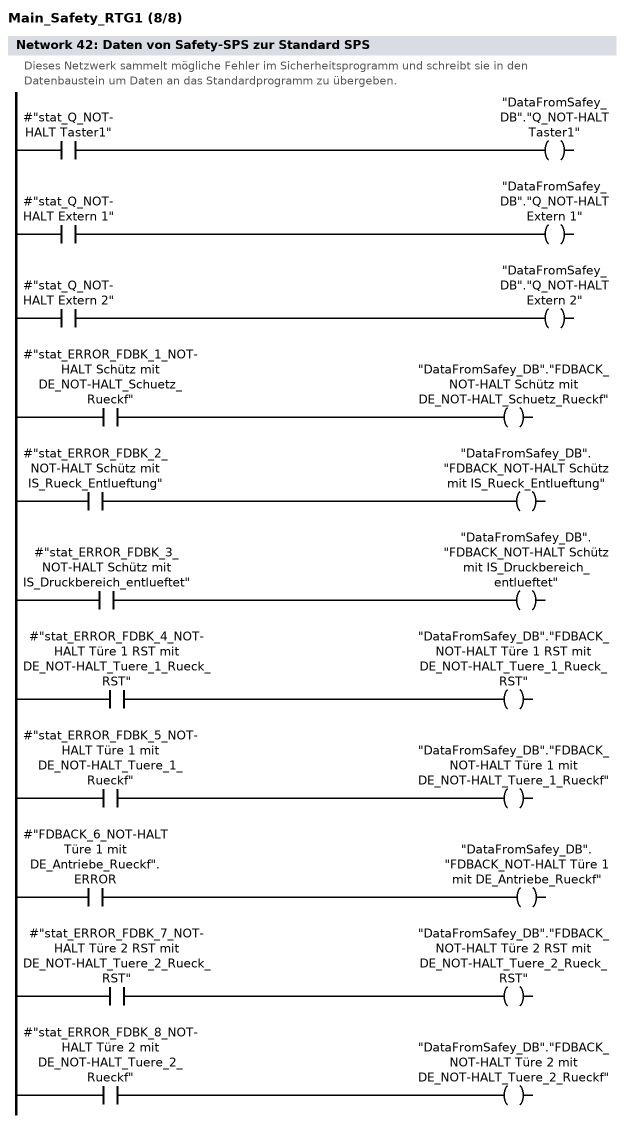
   RUNG wire#powerrail
      Contact( #"stat_Q_NOT-HALT Taster1" )
      Coil( "DataFromSafey_DB"."Q_NOT-HALT Taster1" )
   END_RUNG
   RUNG wire#powerrail
      Contact( #"stat_Q_NOT-HALT Extern 1" )
      Coil( "DataFromSafey_DB"."Q_NOT-HALT Extern 1" )
   END_RUNG
   RUNG wire#powerrail
      Contact( #"stat_Q_NOT-HALT Extern 2" )
      Coil( "DataFromSafey_DB"."Q_NOT-HALT Extern 2" )
   END_RUNG
   RUNG wire#powerrail
      Contact( #"stat_ERROR_FDBK_1_NOT-HALT Schütz mit DE_NOT-HALT_Schuetz_Rueckf" )
      Coil( "DataFromSafey_DB"."FDBACK_NOT-HALT Schütz mit DE_NOT-HALT_Schuetz_Rueckf" )
   END_RUNG
   RUNG wire#powerrail
      Contact( #"stat_ERROR_FDBK_2_NOT-HALT Schütz mit IS_Rueck_Entlueftung" )
      Coil( "DataFromSafey_DB"."FDBACK_NOT-HALT Schütz mit IS_Rueck_Entlueftung" )
   END_RUNG
   RUNG wire#powerrail
      Contact( #"stat_ERROR_FDBK_3_NOT-HALT Schütz mit IS_Druckbereich_entlueftet" )
      Coil( "DataFromSafey_DB"."FDBACK_NOT-HALT Schütz mit IS_Druckbereich_entlueftet" )
   END_RUNG
   RUNG wire#powerrail
      Contact( #"stat_ERROR_FDBK_4_NOT-HALT Türe 1 RST mit DE_NOT-HALT_Tuere_1_Rueck_RST" )
      Coil( "DataFromSafey_DB"."FDBACK_NOT-HALT Türe 1 RST mit DE_NOT-HALT_Tuere_1_Rueck_RST" )
   END_RUNG
   RUNG wire#powerrail
      Contact( #"stat_ERROR_FDBK_5_NOT-HALT Türe 1 mit DE_NOT-HALT_Tuere_1_Rueckf" )
      Coil( "DataFromSafey_DB"."FDBACK_NOT-HALT Türe 1 mit DE_NOT-HALT_Tuere_1_Rueckf" )
   END_RUNG
   RUNG wire#powerrail
      Contact( #"FDBACK_6_NOT-HALT Türe 1 mit DE_Antriebe_Rueckf".ERROR )
      Coil( "DataFromSafey_DB"."FDBACK_NOT-HALT Türe 1 mit DE_Antriebe_Rueckf" )
   END_RUNG
   RUNG wire#powerrail
      Contact( #"stat_ERROR_FDBK_7_NOT-HALT Türe 2 RST mit DE_NOT-HALT_Tuere_2_Rueck_RST" )
      Coil( "DataFromSafey_DB"."FDBACK_NOT-HALT Türe 2 RST mit DE_NOT-HALT_Tuere_2_Rueck_RST" )
   END_RUNG
   RUNG wire#powerrail
      Contact( #"stat_ERROR_FDBK_8_NOT-HALT Türe 2 mit DE_NOT-HALT_Tuere_2_Rueckf" )
      Coil( "DataFromSafey_DB"."FDBACK_NOT-HALT Türe 2 mit DE_NOT-HALT_Tuere_2_Rueckf" )
   END_RUNG
   // the same network as SCL:
   "DataFromSafey_DB"."Q_NOT-HALT Taster1" := #"stat_Q_NOT-HALT Taster1";
   "DataFromSafey_DB"."Q_NOT-HALT Extern 1" := #"stat_Q_NOT-HALT Extern 1";
   "DataFromSafey_DB"."Q_NOT-HALT Extern 2" := #"stat_Q_NOT-HALT Extern 2";
   "DataFromSafey_DB"."FDBACK_NOT-HALT Schütz mit DE_NOT-HALT_Schuetz_Rueckf" := #"stat_ERROR_FDBK_1_NOT-HALT Schütz mit DE_NOT-HALT_Schuetz_Rueckf";
   "DataFromSafey_DB"."FDBACK_NOT-HALT Schütz mit IS_Rueck_Entlueftung" := #"stat_ERROR_FDBK_2_NOT-HALT Schütz mit IS_Rueck_Entlueftung";
   "DataFromSafey_DB"."FDBACK_NOT-HALT Schütz mit IS_Druckbereich_entlueftet" := #"stat_ERROR_FDBK_3_NOT-HALT Schütz mit IS_Druckbereich_entlueftet";
   "DataFromSafey_DB"."FDBACK_NOT-HALT Türe 1 RST mit DE_NOT-HALT_Tuere_1_Rueck_RST" := #"stat_ERROR_FDBK_4_NOT-HALT Türe 1 RST mit DE_NOT-HALT_Tuere_1_Rueck_RST";
   "DataFromSafey_DB"."FDBACK_NOT-HALT Türe 1 mit DE_NOT-HALT_Tuere_1_Rueckf" := #"stat_ERROR_FDBK_5_NOT-HALT Türe 1 mit DE_NOT-HALT_Tuere_1_Rueckf";
   "DataFromSafey_DB"."FDBACK_NOT-HALT Türe 1 mit DE_Antriebe_Rueckf" := #"FDBACK_6_NOT-HALT Türe 1 mit DE_Antriebe_Rueckf".ERROR;
   "DataFromSafey_DB"."FDBACK_NOT-HALT Türe 2 RST mit DE_NOT-HALT_Tuere_2_Rueck_RST" := #"stat_ERROR_FDBK_7_NOT-HALT Türe 2 RST mit DE_NOT-HALT_Tuere_2_Rueck_RST";
   "DataFromSafey_DB"."FDBACK_NOT-HALT Türe 2 mit DE_NOT-HALT_Tuere_2_Rueckf" := #"stat_ERROR_FDBK_8_NOT-HALT Türe 2 mit DE_NOT-HALT_Tuere_2_Rueckf";
END_REGION
END_FUNCTION_BLOCK
